{attribute 'qualified_only'}
{attribute 'strict'}
//{attribute 'to_string'}
TYPE E_MirrorCoverState :
(
	closing := 0,
	opening := 1,
	stopped := 2,
	closed	:= 3,
	open	:= 4,
	error := 5,
	unknown := 6
);
END_TYPE

(* stored: Version 1.1.0.1, ProductVersion 3.1.4024.12
   DUT E_MirrorCoverState: Id {912d241f-d2a8-419d-8f08-9f22cedc1d83} *)
